FUNCTION_BLOCK fbrisetrig
VAR_INPUT
	clkin:BOOL;
	
END_VAR
VAR_OUTPUT
	clkout:BOOL;
	
END_VAR
VAR
	bprevclk:BOOL;
	
END_VAR

clkout:= clkin AND NOT bprevclk;
bprevclk:=clkin;

END_FUNCTION_BLOCK

(* stored: Version 1.1.0.1, ProductVersion 3.1.4024.16
   POU fbrisetrig: Id {eb5d26b5-5673-416e-9bef-f173508a7ffa}, SpecialFunc None *)
